(* IEC 61131-3 sources: plc-process-lib/tests/POUs/Suites/FB_DigitalInput_Test, 28 files *)

(* ---- AlarmEventsValueIsZeroOrOne.method.decl.st ---- *)
// Значение события тревог дискретного входа — xValue как 1.0 / 0.0 (DI-7): State при xValue = TRUE — Activated со
// значением 1.0, снятие — Cleared со значением 0.0; номер тревоги State = udiAlarmIdBase + 0.
METHOD PRIVATE AlarmEventsValueIsZeroOrOne
VAR
    fbTime  : FB_FakeTime;          // подменное время
    fbDi    : FB_DigitalInput;      // ФБ под тестом
    stCmd   : ST_DigitalInputCmd;   // команды
    stCfg   : ST_DigitalInputCfg;   // конфигурация
    fbSink  : FB_TestSink;          // приёмник событий
    stEvOn  : ST_AlarmEvent;        // событие появления
    stEvOff : ST_AlarmEvent;        // событие снятия
END_VAR

(* ---- AlarmOnFalseActivatesWhenValueFalse.method.decl.st ---- *)
// xAlarmOnTrue = FALSE (тревога при пропадании сигнала, например «давление в норме»): TRUE — тревоги нет; FALSE —
// тревога State ActiveUnack, бит DI_STS_ALARM_COND, приоритет в ePrioUnack.
METHOD PRIVATE AlarmOnFalseActivatesWhenValueFalse
VAR
    fbTime : FB_FakeTime;          // подменное время
    fbDi   : FB_DigitalInput;      // ФБ под тестом
    stCmd  : ST_DigitalInputCmd;   // команды
    stCfg  : ST_DigitalInputCfg;   // конфигурация
    itfAlm : I_Alarm;              // слот тревоги через интерфейс
END_VAR

(* ---- ChannelFaultDuringOnDelayRestartsDelay.method.decl.st ---- *)
// Отказ канала во время задержки включения: сигнал при отказе недостоверен, поэтому задержка после возврата канала
// отсчитывается заново (DI-2), а не продолжается с момента фронта; биты отсчёта во время отказа не выставляются.
// tOnDelay = 1 с: фронт в t0, отказ t0 + 0,6 … t0 + 0,8 с, возврат tr = t0 + 0,8 с — значение в tr + 1,0 с.
METHOD PRIVATE ChannelFaultDuringOnDelayRestartsDelay
VAR
    fbTime  : FB_FakeTime;          // подменное время
    fbDi    : FB_DigitalInput;      // ФБ под тестом
    stCmd   : ST_DigitalInputCmd;   // команды
    stCfg   : ST_DigitalInputCfg;   // конфигурация
    iStep   : INT;                  // шаг цикла
    xEverOn : BOOL;                 // значение включалось хотя бы раз
END_VAR

(* ---- ChannelFaultDuringOnDelayRestartsDelay.method.impl.st ---- *)
coUnit.TEST('DigitalInput_ChannelFaultDuringOnDelay_RestartsDelay');

stCfg.tOnDelay := T#1S;
fbDi(itfTime := fbTime, xIn := FALSE, stCmd := stCmd, stCfg := stCfg);
fbTime.Advance(tStep := T#100MS);
fbDi(itfTime := fbTime, xIn := TRUE, stCmd := stCmd, stCfg := stCfg);   // t0: фронт
FOR iStep := 1 TO 5 DO   // t0 + 0,5 с
    fbTime.Advance(tStep := T#100MS);
    fbDi(itfTime := fbTime, xIn := TRUE, stCmd := stCmd, stCfg := stCfg);
END_FOR
AssertTrue(Condition := (fbDi.stSts.stCommon.wStatus AND GVL_Const.DI_STS_TIMING_ON) <> 0, Message := 'timing on');
FOR iStep := 1 TO 2 DO   // отказ канала: t0 + 0,6 … t0 + 0,7 с
    fbTime.Advance(tStep := T#100MS);
    fbDi(itfTime := fbTime, xIn := TRUE, xChannelFault := TRUE, stCmd := stCmd, stCfg := stCfg);
END_FOR
AssertTrue(Condition := (fbDi.stSts.stCommon.wStatus AND GVL_Const.DI_STS_TIMING_ON) = 0,
           Message := 'no timing bit during channel fault');
AssertFalse(Condition := fbDi.xValue, Message := 'value before the fault held');
fbTime.Advance(tStep := T#100MS);
fbDi(itfTime := fbTime, xIn := TRUE, xChannelFault := FALSE, stCmd := stCmd, stCfg := stCfg);   // tr = t0 + 0,8 с
xEverOn := fbDi.xValue;
FOR iStep := 1 TO 9 DO   // tr + 0,9 с (t0 + 1,7 с)
    fbTime.Advance(tStep := T#100MS);
    fbDi(itfTime := fbTime, xIn := TRUE, stCmd := stCmd, stCfg := stCfg);
    xEverOn := xEverOn OR fbDi.xValue;
END_FOR
AssertFalse(Condition := xEverOn, Message := 'on-delay restarted at recovery, not counted from t0');
AssertTrue(Condition := (fbDi.stSts.stCommon.wStatus AND GVL_Const.DI_STS_TIMING_ON) <> 0,
           Message := 'timing on again after recovery');
fbTime.Advance(tStep := T#100MS);
fbDi(itfTime := fbTime, xIn := TRUE, stCmd := stCmd, stCfg := stCfg);   // tr + 1,0 с
AssertTrue(Condition := fbDi.xValue, Message := 'value exactly tOnDelay after recovery');

coUnit.TEST_FINISHED();

(* ---- ChannelFaultForceFalse.method.decl.st ---- *)
// ForceFalse: отказ канала при включённом сигнале — значение FALSE сразу, xValid = FALSE.
METHOD PRIVATE ChannelFaultForceFalse
VAR
    fbTime : FB_FakeTime;          // подменное время
    fbDi   : FB_DigitalInput;      // ФБ под тестом
    stCmd  : ST_DigitalInputCmd;   // команды
    stCfg  : ST_DigitalInputCfg;   // конфигурация
END_VAR

(* ---- ChannelFaultForceTrue.method.decl.st ---- *)
// ForceTrue (защитный сигнал: отказ канала = сработал): отказ — значение TRUE сразу, xValid = FALSE, Failure, биты
// DI_FLT_CHANNEL и DI_STS_CHANNEL_FAULT, тревога Failure ActiveUnack, тревога State подавлена (SuppressedByDesign, без
// дублирования). Отказ снят — снова измерение.
METHOD PRIVATE ChannelFaultForceTrue
VAR
    fbTime : FB_FakeTime;          // подменное время
    fbDi   : FB_DigitalInput;      // ФБ под тестом
    stCmd  : ST_DigitalInputCmd;   // команды
    stCfg  : ST_DigitalInputCfg;   // конфигурация
    itfAlm : I_Alarm;              // слот тревоги через интерфейс
END_VAR

(* ---- ChannelFaultHoldLast.method.decl.st ---- *)
// HoldLast: при отказе канала держится значение до отказа (TRUE), xValid = FALSE; после отказа задержка отключения 1 с
// отсчитывается от возврата канала.
METHOD PRIVATE ChannelFaultHoldLast
VAR
    fbTime : FB_FakeTime;          // подменное время
    fbDi   : FB_DigitalInput;      // ФБ под тестом
    stCmd  : ST_DigitalInputCmd;   // команды
    stCfg  : ST_DigitalInputCfg;   // конфигурация
    iStep  : INT;                  // шаг цикла
END_VAR

(* ---- ChannelFaultHoldLast.method.impl.st ---- *)
coUnit.TEST('DigitalInput_ChannelFault_HoldLast');

stCfg.tOffDelay := T#1S;
fbDi(itfTime := fbTime, xIn := TRUE, stCmd := stCmd, stCfg := stCfg);
FOR iStep := 1 TO 5 DO   // отказ канала 0,5 с
    fbTime.Advance(tStep := T#100MS);
    fbDi(itfTime := fbTime, xIn := FALSE, xChannelFault := TRUE, stCmd := stCmd, stCfg := stCfg);
END_FOR
AssertTrue(Condition := fbDi.xValue, Message := 'value before the fault held');
AssertFalse(Condition := fbDi.xValid, Message := 'invalid during fault');
fbTime.Advance(tStep := T#100MS);
fbDi(itfTime := fbTime, xIn := FALSE, xChannelFault := FALSE, stCmd := stCmd, stCfg := stCfg);   // tr: канал исправен
AssertTrue(Condition := fbDi.xValue, Message := 'off-delay restarts at recovery');
AssertTrue(Condition := fbDi.xValid, Message := 'valid after recovery');
FOR iStep := 1 TO 9 DO   // tr + 0,9 с
    fbTime.Advance(tStep := T#100MS);
    fbDi(itfTime := fbTime, xIn := FALSE, xChannelFault := FALSE, stCmd := stCmd, stCfg := stCfg);
END_FOR
AssertTrue(Condition := fbDi.xValue, Message := 'held until tr + 1.0 s');
fbTime.Advance(tStep := T#100MS);
fbDi(itfTime := fbTime, xIn := FALSE, xChannelFault := FALSE, stCmd := stCmd, stCfg := stCfg);   // tr + 1,0 с
AssertFalse(Condition := fbDi.xValue, Message := 'off after off-delay from recovery');

coUnit.TEST_FINISHED();

(* ---- ChannelFaultRecoveredForcedValueReleasedThroughDelay.method.decl.st ---- *)
// Защитный сигнал (ForceTrue, «сухой ход»): после возврата канала задержки отсчитываются от значения отказа, а не
// от значения до отказа (DI-2). tOnDelay 2 с, tOffDelay 3 с. 1) До отказа FALSE, после возврата датчик сработал
// (TRUE) — значение остаётся TRUE без провала (иначе 2 с FALSE при xValid = TRUE: насос пустили бы на сухую).
// 2) До отказа FALSE, после возврата датчик в норме — TRUE снимается только через tOffDelay, ровно в tr + 3,0 с.
METHOD PRIVATE ChannelFaultRecoveredForcedValueReleasedThroughDelay
VAR
    fbTime   : FB_FakeTime;          // подменное время
    fbDi     : FB_DigitalInput;      // ФБ под тестом
    stCmd    : ST_DigitalInputCmd;   // команды
    stCfg    : ST_DigitalInputCfg;   // конфигурация
    iStep    : INT;                  // шаг цикла
    xEverOff : BOOL;                 // значение выключалось хотя бы раз
END_VAR

(* ---- ChannelFaultRecoveredForcedValueReleasedThroughDelay.method.impl.st ---- *)
coUnit.TEST('DigitalInput_ChannelFaultRecovered_ForcedValueReleasedThroughDelay');

stCfg.eFailValue := E_DiFailValue.ForceTrue;
stCfg.tOnDelay := T#2S;
stCfg.tOffDelay := T#3S;
fbDi(itfTime := fbTime, xIn := FALSE, stCmd := stCmd, stCfg := stCfg);   // норма: FALSE
fbTime.Advance(tStep := T#100MS);
fbDi(itfTime := fbTime, xIn := FALSE, xChannelFault := TRUE, stCmd := stCmd, stCfg := stCfg);   // отказ канала
AssertTrue(Condition := fbDi.xValue, Message := 'forced TRUE on channel fault');
// 1) канал исправен, датчик сработал
fbTime.Advance(tStep := T#100MS);
fbDi(itfTime := fbTime, xIn := TRUE, xChannelFault := FALSE, stCmd := stCmd, stCfg := stCfg);
xEverOff := NOT fbDi.xValue;
AssertTrue(Condition := fbDi.xValid, Message := 'valid after recovery');
FOR iStep := 1 TO 25 DO   // 2,5 с: дольше tOnDelay
    fbTime.Advance(tStep := T#100MS);
    fbDi(itfTime := fbTime, xIn := TRUE, stCmd := stCmd, stCfg := stCfg);
    xEverOff := xEverOff OR NOT fbDi.xValue;
END_FOR
AssertFalse(Condition := xEverOff, Message := 'no FALSE gap after recovery when the sensor is tripped');
// 2) датчик в норме дольше tOffDelay, затем отказ и возврат с датчиком в норме
FOR iStep := 1 TO 31 DO   // 3,1 с
    fbTime.Advance(tStep := T#100MS);
    fbDi(itfTime := fbTime, xIn := FALSE, stCmd := stCmd, stCfg := stCfg);
END_FOR
AssertFalse(Condition := fbDi.xValue, Message := 'value off before the second fault');
fbTime.Advance(tStep := T#100MS);
fbDi(itfTime := fbTime, xIn := FALSE, xChannelFault := TRUE, stCmd := stCmd, stCfg := stCfg);
fbTime.Advance(tStep := T#100MS);
fbDi(itfTime := fbTime, xIn := FALSE, xChannelFault := FALSE, stCmd := stCmd, stCfg := stCfg);   // tr: канал исправен
AssertTrue(Condition := fbDi.xValue, Message := 'forced value kept at recovery');
FOR iStep := 1 TO 29 DO   // tr + 2,9 с
    fbTime.Advance(tStep := T#100MS);
    fbDi(itfTime := fbTime, xIn := FALSE, stCmd := stCmd, stCfg := stCfg);
END_FOR
AssertTrue(Condition := fbDi.xValue, Message := 'released only through tOffDelay');
AssertTrue(Condition := (fbDi.stSts.stCommon.wStatus AND GVL_Const.DI_STS_TIMING_OFF) <> 0, Message := 'timing off');
fbTime.Advance(tStep := T#100MS);
fbDi(itfTime := fbTime, xIn := FALSE, stCmd := stCmd, stCfg := stCfg);   // tr + 3,0 с
AssertFalse(Condition := fbDi.xValue, Message := 'off exactly tOffDelay after recovery');

coUnit.TEST_FINISHED();

(* ---- DefaultCfgFirstCallValueWithoutDelay.method.decl.st ---- *)
// Cfg по умолчанию проходит CheckConfig; после первого вызова — Auto, тип DigitalInput, 2 слота, Good. Значение в
// первом вызове — без задержки включения (2 с): после старта ПЛК вход сразу равен сигналу. Тревога State по умолчанию
// выключена (None) и не формируется.
METHOD PRIVATE DefaultCfgFirstCallValueWithoutDelay
VAR
    fbTime : FB_FakeTime;          // подменное время
    fbDi   : FB_DigitalInput;      // ФБ под тестом
    stCmd  : ST_DigitalInputCmd;   // команды
    stCfg  : ST_DigitalInputCfg;   // конфигурация
    itfAlm : I_Alarm;              // слот тревоги через интерфейс
END_VAR

(* ---- InvalidCfgAtStartupValueFalseCheckFunction.method.decl.st ---- *)
// Без корректной Cfg с первого вызова (eFailValue и приоритет тревоги вне перечисления): биты DI_CFG_FAIL_VALUE и
// DI_CFG_ALARM, значение FALSE при xIn = TRUE, xValid = FALSE, Available = FALSE, CheckFunction. Исправленная Cfg —
// измерение.
METHOD PRIVATE InvalidCfgAtStartupValueFalseCheckFunction
VAR
    fbTime : FB_FakeTime;          // подменное время
    fbDi   : FB_DigitalInput;      // ФБ под тестом
    stCmd  : ST_DigitalInputCmd;   // команды
    stCfg  : ST_DigitalInputCfg;   // конфигурация
    uEnum  : U_AiDiTestEnum;       // значение вне строгого перечисления
    uPrio  : U_TestEnumInt;        // приоритет вне перечисления
END_VAR

(* ---- InvertFromFirstValidCfgNoFalseValue.method.decl.st ---- *)
// Корректная Cfg появилась не в первом вызове (на старте Cfg была испорчена, наладчик исправил её с HMI): задержки
// предустанавливаются по сигналу с инверсией из этой Cfg, а не по сигналу без инверсии, который считался по
// умолчаниям Cfg. Поплавок «сухой ход», НЗ-контакт (xInvert), задержки 2 с: A — контакт замкнут (норма) — значение
// FALSE сразу, без ложного «сухого хода» на tOffDelay; B — контакт разомкнут (сработал) — TRUE сразу, без пропуска
// срабатывания на tOnDelay.
METHOD PRIVATE InvertFromFirstValidCfgNoFalseValue
VAR
    fbTime : FB_FakeTime;          // подменное время
    fbDiA  : FB_DigitalInput;      // контакт замкнут
    fbDiB  : FB_DigitalInput;      // контакт разомкнут
    stCmdA : ST_DigitalInputCmd;   // команды A
    stCmdB : ST_DigitalInputCmd;   // команды B
    stCfg  : ST_DigitalInputCfg;   // конфигурация
    uEnum  : U_AiDiTestEnum;       // значение вне строгого перечисления
END_VAR

(* ---- InvertInvertsBeforeDelay.method.decl.st ---- *)
// Инверсия (НЗ-контакт) до задержек: xIn TRUE — значение FALSE; пропадание xIn — фронт инвертированного сигнала, его и
// задерживает tOnDelay 300 мс (бит DI_STS_RAW = 1 сразу); возврат xIn — спад без задержки.
METHOD PRIVATE InvertInvertsBeforeDelay
VAR
    fbTime : FB_FakeTime;          // подменное время
    fbDi   : FB_DigitalInput;      // ФБ под тестом
    stCmd  : ST_DigitalInputCmd;   // команды
    stCfg  : ST_DigitalInputCfg;   // конфигурация
    iStep  : INT;                  // шаг цикла
END_VAR

(* ---- InvertInvertsBeforeDelay.method.impl.st ---- *)
coUnit.TEST('DigitalInput_Invert_InvertsBeforeDelay');

stCfg.xInvert := TRUE;
stCfg.tOnDelay := T#300MS;
fbDi(itfTime := fbTime, xIn := TRUE, stCmd := stCmd, stCfg := stCfg);   // t0
AssertFalse(Condition := fbDi.xValue, Message := 'inverted: TRUE gives FALSE');
AssertTrue(Condition := (fbDi.stSts.stCommon.wStatus AND GVL_Const.DI_STS_RAW) = 0, Message := 'raw after inversion');
fbTime.Advance(tStep := T#100MS);
fbDi(itfTime := fbTime, xIn := FALSE, stCmd := stCmd, stCfg := stCfg);   // t1: разрыв НЗ-контакта
AssertTrue(Condition := (fbDi.stSts.stCommon.wStatus AND GVL_Const.DI_STS_RAW) <> 0, Message := 'raw TRUE at once');
FOR iStep := 1 TO 2 DO   // t1 + 0,2 с
    fbTime.Advance(tStep := T#100MS);
    fbDi(itfTime := fbTime, xIn := FALSE, stCmd := stCmd, stCfg := stCfg);
END_FOR
AssertFalse(Condition := fbDi.xValue, Message := 'on-delay applies to the inverted signal');
fbTime.Advance(tStep := T#100MS);
fbDi(itfTime := fbTime, xIn := FALSE, stCmd := stCmd, stCfg := stCfg);   // t1 + 0,3 с
AssertTrue(Condition := fbDi.xValue, Message := 'value after on-delay');
fbTime.Advance(tStep := T#100MS);
fbDi(itfTime := fbTime, xIn := TRUE, stCmd := stCmd, stCfg := stCfg);
AssertFalse(Condition := fbDi.xValue, Message := 'falling edge without off-delay');

coUnit.TEST_FINISHED();

(* ---- OffDelayHoldsValue.method.decl.st ---- *)
// Задержка отключения 1 с: сигнал пропал — значение держится 0,9 с (бит DI_STS_TIMING_OFF), снимается ровно через 1,0
// с.
METHOD PRIVATE OffDelayHoldsValue
VAR
    fbTime : FB_FakeTime;          // подменное время
    fbDi   : FB_DigitalInput;      // ФБ под тестом
    stCmd  : ST_DigitalInputCmd;   // команды
    stCfg  : ST_DigitalInputCfg;   // конфигурация
    iStep  : INT;                  // шаг цикла
END_VAR

(* ---- OffDelayHoldsValue.method.impl.st ---- *)
coUnit.TEST('DigitalInput_OffDelay_HoldsValue');

stCfg.tOffDelay := T#1S;
fbDi(itfTime := fbTime, xIn := TRUE, stCmd := stCmd, stCfg := stCfg);   // t0
AssertTrue(Condition := fbDi.xValue, Message := 'value on');
fbTime.Advance(tStep := T#100MS);
fbDi(itfTime := fbTime, xIn := FALSE, stCmd := stCmd, stCfg := stCfg);   // t1: сигнал пропал
FOR iStep := 1 TO 9 DO   // t1 + 0,9 с
    fbTime.Advance(tStep := T#100MS);
    fbDi(itfTime := fbTime, xIn := FALSE, stCmd := stCmd, stCfg := stCfg);
END_FOR
AssertTrue(Condition := fbDi.xValue, Message := 'value held by off-delay');
AssertTrue(Condition := (fbDi.stSts.stCommon.wStatus AND GVL_Const.DI_STS_TIMING_OFF) <> 0,
           Message := 'timing off bit');
fbTime.Advance(tStep := T#100MS);
fbDi(itfTime := fbTime, xIn := FALSE, stCmd := stCmd, stCfg := stCfg);   // t1 + 1,0 с
AssertFalse(Condition := fbDi.xValue, Message := 'value off after off-delay');

coUnit.TEST_FINISHED();

(* ---- OnDelayFiltersBounce.method.decl.st ---- *)
// Задержка включения 500 мс: дребезг (импульсы 200 и 300 мс) значение не включает, пока идёт отсчёт — бит
// DI_STS_TIMING_ON; устойчивый сигнал — TRUE ровно через 500 мс.
METHOD PRIVATE OnDelayFiltersBounce
VAR
    fbTime  : FB_FakeTime;          // подменное время
    fbDi    : FB_DigitalInput;      // ФБ под тестом
    stCmd   : ST_DigitalInputCmd;   // команды
    stCfg   : ST_DigitalInputCfg;   // конфигурация
    iStep   : INT;                  // шаг цикла
    xEverOn : BOOL;                 // значение включалось хотя бы раз
END_VAR

(* ---- OnDelayFiltersBounce.method.impl.st ---- *)
coUnit.TEST('DigitalInput_OnDelay_FiltersBounce');

stCfg.tOnDelay := T#500MS;
fbDi(itfTime := fbTime, xIn := FALSE, stCmd := stCmd, stCfg := stCfg);   // t0
FOR iStep := 1 TO 2 DO                                            // импульс 200 мс
    fbTime.Advance(tStep := T#100MS);
    fbDi(itfTime := fbTime, xIn := TRUE, stCmd := stCmd, stCfg := stCfg);
    xEverOn := xEverOn OR fbDi.xValue;
END_FOR
AssertTrue(Condition := (fbDi.stSts.stCommon.wStatus AND GVL_Const.DI_STS_TIMING_ON) <> 0, Message := 'timing on bit');
AssertTrue(Condition := (fbDi.stSts.stCommon.wStatus AND GVL_Const.DI_STS_RAW) <> 0, Message := 'raw bit');
fbTime.Advance(tStep := T#100MS);
fbDi(itfTime := fbTime, xIn := FALSE, stCmd := stCmd, stCfg := stCfg);
FOR iStep := 1 TO 3 DO                                            // импульс 300 мс
    fbTime.Advance(tStep := T#100MS);
    fbDi(itfTime := fbTime, xIn := TRUE, stCmd := stCmd, stCfg := stCfg);
    xEverOn := xEverOn OR fbDi.xValue;
END_FOR
fbTime.Advance(tStep := T#100MS);
fbDi(itfTime := fbTime, xIn := FALSE, stCmd := stCmd, stCfg := stCfg);
xEverOn := xEverOn OR fbDi.xValue;
AssertFalse(Condition := xEverOn, Message := 'bounce shorter than on-delay ignored');
fbTime.Advance(tStep := T#100MS);
fbDi(itfTime := fbTime, xIn := TRUE, stCmd := stCmd, stCfg := stCfg);   // t1: устойчивый сигнал
FOR iStep := 1 TO 4 DO   // t1 + 0,4 с
    fbTime.Advance(tStep := T#100MS);
    fbDi(itfTime := fbTime, xIn := TRUE, stCmd := stCmd, stCfg := stCfg);
END_FOR
AssertFalse(Condition := fbDi.xValue, Message := 'no value at t1 + 0.4 s');
fbTime.Advance(tStep := T#100MS);
fbDi(itfTime := fbTime, xIn := TRUE, stCmd := stCmd, stCfg := stCfg);   // t1 + 0,5 с
AssertTrue(Condition := fbDi.xValue, Message := 'value exactly at t1 + 0.5 s');
AssertTrue(Condition := (fbDi.stSts.stCommon.wStatus AND GVL_Const.DI_STS_VALUE) <> 0, Message := 'value bit');
AssertTrue(Condition := (fbDi.stSts.stCommon.wStatus AND GVL_Const.DI_STS_TIMING_ON) = 0, Message := 'timing done');

coUnit.TEST_FINISHED();

(* ---- OutOfServiceAlarmsOutOfService.method.decl.st ---- *)
// OutOfService: оба слота OutOfService (в wAlmShelved их нет — ALM-2), значение удерживается (TRUE), xValid = FALSE,
// CheckFunction; отказ канала в OOS не даёт Failure; слежение xSubstValue действует и в OOS (2.1). После выхода
// активная тревога State снова ActiveUnack.
METHOD PRIVATE OutOfServiceAlarmsOutOfService
VAR
    fbTime : FB_FakeTime;          // подменное время
    fbDi   : FB_DigitalInput;      // ФБ под тестом
    stCmd  : ST_DigitalInputCmd;   // команды
    stCfg  : ST_DigitalInputCfg;   // конфигурация
    itfAlm : I_Alarm;              // слот тревоги через интерфейс
END_VAR

(* ---- ResetCmdAcceptedAndAcksAlarms.method.decl.st ---- *)
// xReset у DI — команда без фиксируемых отказов: результат Accepted, uiCmdSeq + 1, бит сброшен; тревога Failure после
// отказа канала (RtnUnack) квитирована.
METHOD PRIVATE ResetCmdAcceptedAndAcksAlarms
VAR
    fbTime : FB_FakeTime;          // подменное время
    fbDi   : FB_DigitalInput;      // ФБ под тестом
    stCmd  : ST_DigitalInputCmd;   // команды
    stCfg  : ST_DigitalInputCfg;   // конфигурация
    itfAlm : I_Alarm;              // слот тревоги через интерфейс
    uiSeq  : UINT;                 // номер команды до сброса
END_VAR

(* ---- SetAlarmPriority.method.decl.st ---- *)
// Помощник: приоритет слота тревоги uiSlot в Cfg входа (через копию элемента)
METHOD PRIVATE SetAlarmPriority
VAR_IN_OUT
    stCfgDi : ST_DigitalInputCfg;  // конфигурация входа
END_VAR
VAR_INPUT
    uiSlot    : UINT;              // слот: E_DiAlarm
    ePriority : E_AlarmPriority;   // приоритет
END_VAR
VAR
    stSlot : ST_AlarmCfg;          // копия слота
END_VAR

(* ---- SubstitutionOverridesValueBypassesDelay.method.decl.st ---- *)
// Подмена (Manual): значение — stCmd.xSubstValue в том же вызове, без задержек 5 с; пригодно, NE 107 CheckFunction. До
// подмены ФБ следит: stCmd.xSubstValue = xValue.
METHOD PRIVATE SubstitutionOverridesValueBypassesDelay
VAR
    fbTime : FB_FakeTime;          // подменное время
    fbDi   : FB_DigitalInput;      // ФБ под тестом
    stCmd  : ST_DigitalInputCmd;   // команды
    stCfg  : ST_DigitalInputCfg;   // конфигурация
END_VAR

(* ---- SubstitutionRenewedAfterTimeoutCountsFullPeriod.method.decl.st ---- *)
// Подмена, снятая по tSubstMax, и новый запрос подмены в следующем же вызове: срок отсчитывается заново, подмена не
// снимается сразу же. Остаток uiSubstRemain_s — целые секунды с округлением вверх (29,4 с -> 30, 0,3 с -> 1).
METHOD PRIVATE SubstitutionRenewedAfterTimeoutCountsFullPeriod
VAR
    fbTime : FB_FakeTime;          // подменное время
    fbDi   : FB_DigitalInput;      // ФБ под тестом
    stCmd  : ST_DigitalInputCmd;   // команды
    stCfg  : ST_DigitalInputCfg;   // конфигурация
END_VAR

(* ---- SubstitutionTimeoutReturnsToAuto.method.decl.st ---- *)
// tSubstMax 30 с: подмена TRUE; остаток 30 при входе, 1 в 29 с; ровно через 30 с — Auto, результат SubstExpired,
// значение измеренное (FALSE).
METHOD PRIVATE SubstitutionTimeoutReturnsToAuto
VAR
    fbTime : FB_FakeTime;          // подменное время
    fbDi   : FB_DigitalInput;      // ФБ под тестом
    stCmd  : ST_DigitalInputCmd;   // команды
    stCfg  : ST_DigitalInputCfg;   // конфигурация
    iStep  : INT;                  // шаг цикла
END_VAR

(* ---- SubstitutionTimeoutReturnsToAuto.method.impl.st ---- *)
coUnit.TEST('DigitalInput_SubstitutionTimeout_ReturnsToAuto');

stCfg.tSubstMax := T#30S;
fbDi(itfTime := fbTime, xIn := FALSE, stCmd := stCmd, stCfg := stCfg);
stCmd.stCommon.xSetManual := TRUE;
stCmd.xSubstValue := TRUE;
fbTime.Advance(tStep := T#100MS);
fbDi(itfTime := fbTime, xIn := FALSE, stCmd := stCmd, stCfg := stCfg);   // t0: подмена
AssertEquals_UINT(Expected := 30, Actual := fbDi.stSts.uiSubstRemain_s, Message := '30 s remain at start');
FOR iStep := 1 TO 29 DO   // t0 + 29 с
    fbTime.Advance(tStep := T#1000MS);
    fbDi(itfTime := fbTime, xIn := FALSE, stCmd := stCmd, stCfg := stCfg);
END_FOR
AssertTrue(Condition := fbDi.Mode = E_DeviceMode.Manual, Message := 'still substituted');
AssertTrue(Condition := fbDi.xValue, Message := 'substituted TRUE');
AssertEquals_UINT(Expected := 1, Actual := fbDi.stSts.uiSubstRemain_s, Message := '1 s remains');
fbTime.Advance(tStep := T#1000MS);
fbDi(itfTime := fbTime, xIn := FALSE, stCmd := stCmd, stCfg := stCfg);   // t0 + 30 с
AssertTrue(Condition := fbDi.Mode = E_DeviceMode.Auto, Message := 'back to measurement');
AssertTrue(Condition := fbDi.stSts.stCommon.eCmdResult = E_CmdResult.SubstExpired, Message := 'SubstExpired');
AssertFalse(Condition := fbDi.xValue, Message := 'measured value');
AssertEquals_UINT(Expected := 0, Actual := fbDi.stSts.uiSubstRemain_s, Message := 'no remaining time');

coUnit.TEST_FINISHED();

(* ---- SubstitutionUnlimitedNoTimeout.method.decl.st ---- *)
// tSubstMax = T#0S — подмена без ограничения срока: 24 ч в Manual — режим Manual, SubstExpired нет, значение
// подмены TRUE, остаток 0.
METHOD PRIVATE SubstitutionUnlimitedNoTimeout
VAR
    fbTime    : FB_FakeTime;          // подменное время
    fbDi      : FB_DigitalInput;      // ФБ под тестом
    stCmd     : ST_DigitalInputCmd;   // команды
    stCfg     : ST_DigitalInputCfg;   // конфигурация
    iStep     : INT;                  // шаг цикла
    xEverAuto : BOOL;                 // режим хоть раз вернулся в Auto
END_VAR

(* ---- SubstitutionUnlimitedNoTimeout.method.impl.st ---- *)
coUnit.TEST('DigitalInput_SubstitutionUnlimited_NoTimeout');

stCfg.tSubstMax := T#0S;
fbDi(itfTime := fbTime, xIn := FALSE, stCmd := stCmd, stCfg := stCfg);
stCmd.stCommon.xSetManual := TRUE;
stCmd.xSubstValue := TRUE;
fbTime.Advance(tStep := T#100MS);
fbDi(itfTime := fbTime, xIn := FALSE, stCmd := stCmd, stCfg := stCfg);                 // подмена
AssertTrue(Condition := fbDi.Mode = E_DeviceMode.Manual, Message := 'substituted');
FOR iStep := 1 TO 24 DO
    fbTime.Advance(tStep := T#1H);
    fbDi(itfTime := fbTime, xIn := FALSE, stCmd := stCmd, stCfg := stCfg);
    xEverAuto := xEverAuto OR fbDi.Mode = E_DeviceMode.Auto;
END_FOR
AssertFalse(Condition := xEverAuto, Message := 'never returned to Auto in 24 h');
AssertTrue(Condition := fbDi.stSts.stCommon.eCmdResult = E_CmdResult.Accepted, Message := 'no SubstExpired');
AssertTrue(Condition := fbDi.xValue, Message := 'substituted TRUE');
AssertEquals_UINT(Expected := 0, Actual := fbDi.stSts.uiSubstRemain_s, Message := 'no remaining time without a limit');

coUnit.TEST_FINISHED();
